// TIA Portal V20 export
Screen "Pop-up_PRODDATA_SC_LEGEND_Popup"  340x285
  ScreenItem "Background" at 0,0 size 340x285  Type=HmiRectangle
  ScreenItem "Textfeld_Legende" at 1,1 size 328x25  Type=HmiTextBox
  ScreenItem "Textfeld_11" at 70,196 size 255x89  Type=HmiTextBox
  ScreenItem "Textfeld_8" at 10,238 size 55x30  Type=HmiTextBox
  ScreenItem "Textfeld_9" at 23,219 size 30x20  Type=HmiTextBox
  ScreenItem "Textfeld_13" at 10,190 size 55x30  Type=HmiTextBox
  ScreenItem "Textfeld_10" at 10,34 size 208x28  Type=HmiTextBox
  ScreenItem "Textfeld_14" at 10,63 size 315x35  Type=HmiTextBox
  ScreenItem "Textfeld_2" at 10,100 size 55x30  Type=HmiTextBox
  ScreenItem "Textfeld_3" at 70,100 size 270x96  Type=HmiTextBox
  ScreenItem "Textfeld_4" at 10,133 size 55x30  Type=HmiTextBox
  ScreenItem "Cancel Mode" at 249,3 size 90x60  Type=HmiButton
